Fanuc KAREL source: KB00019.KL

PROGRAM KB00019
%NOLOCKGROUP
%ENVIRONMENT FDEV
VAR
  P1: STRING[80]
  P2: INTEGER
BEGIN
  P1 = 'A'
  P2 = 1
  CHECK_NAME(P1, P2)
END KB00019
